(* IEC 61131-3 sources: JingjiangMoonbox/Application/Application/任务列表/Main_Task/IO配置表_1/KESAI1, 7 files *)

(* ---- KS_AbsEncModule_IODeal_KS1.st ---- *)
(*@CES
Name=KS_AbsEncModule_IODeal_KS1
Type=FunctionBlock
TypeGuid=6f9dac99-8de1-4efc-8465-68ac443b7d08
Guid=41d52946-2a11-4c79-a8c5-b68088c6a3a7
HasDeclaration=True
HasImplementation=False
*)
{DECLARATION}
FUNCTION_BLOCK KS_AbsEncModule_IODeal_KS1
VAR_INPUT
	i_xInputEn:BOOL;
	i_xOutPutEn:BOOL;
	(*这些值的处理未考虑双收双放*)
	i_pdwAbsEncSinglePos_Uw:POINTER TO DWORD;
	i_pwAbsEncMultiPos_Uw:POINTER TO WORD;
	(*收料*)
	i_pdwAbsEncSinglePos_Rw:POINTER TO DWORD;
	i_pwAbsEncMultiPos_Rw:POINTER TO WORD;
	//2025.08.20.152113+
	i_pstStAbsEncIOModule_Uw:POINTER TO StAbsEncIOModule;
	i_pstStAbsEncIOModule_Rw:POINTER TO StAbsEncIOModule;

END_VAR
VAR
	wIWTest:WORD;
	wQWTest: WORD;
	byAbsEncSts: BOOL;
END_VAR

{IMPLEMENTATION}

(* ---- KS_FB_IOMAP_AIAO_KS1.st ---- *)
(*@CES
Name=KS_FB_IOMAP_AIAO_KS1
Type=FunctionBlock
TypeGuid=6f9dac99-8de1-4efc-8465-68ac443b7d08
Guid=356f4cce-85a0-44c7-ab1e-a67fad378d86
HasDeclaration=True
HasImplementation=False
*)
{DECLARATION}
FUNCTION_BLOCK KS_FB_IOMAP_AIAO_KS1
VAR_INPUT
	i_xEn: BOOL;(*功能块使能|*)
	i_xRdInput: BOOL;(*读io输入|*)
	i_xWrOutput: BOOL;(*写io输出|*)
	i_pstStSysParam								: POINTER TO StSysParam;
	i_pastStProgMonitoring						: POINTER TO ARRAY [1..2] OF StProgMonitoring;
END_VAR
VAR_OUTPUT
	o_xEno: BOOL;(*indicated to i_xEn|*)
	o_iErNo: INT;(*0.no err\-1.bad parameter|*)
END_VAR
VAR
//	fb_KS_FB_SetAIType: KS_FB_SetAIType;
	fbKS_FB_Analog_IO_CTL: KS_FB_Analog_IO_CTL;

	byAiFilterTms_UwRw_I					:  BYTE:= 1;(*滤波次数*)
	byAiFilterTms_UwRw_II					:  BYTE:= 1;
	byAiFilterTms_IfOf_I					:  BYTE:= 1;
	byAiFilterTms_IfOf_II					:  BYTE:= 1;
	byAiFilterTms_DiaMeasure_I				:   BYTE:= 1;
	byAiFilterTms_DiaMeasure_II				:   BYTE:= 1;
END_VAR

{IMPLEMENTATION}

(* ---- KS_FB_IOMAP_Axis_KS1.st ---- *)
(*@CES
Name=KS_FB_IOMAP_Axis_KS1
Type=FunctionBlock
TypeGuid=6f9dac99-8de1-4efc-8465-68ac443b7d08
Guid=5e1ef807-2a8d-4def-8e48-4f55f608734d
HasDeclaration=True
HasImplementation=False
*)
{DECLARATION}
FUNCTION_BLOCK KS_FB_IOMAP_Axis_KS1
VAR_INPUT
	i_xEn: BOOL;(*功能块使能|*)
	i_xRdInput: BOOL;(*读io输入|*)
	i_xWrOutput: BOOL;(*写io输出|*)
	i_pastStIOMap_Axis_FE						: POINTER TO ARRAY [1..MAX_UNIT_NUM] OF StIOMap_Axis_FE;(*轴io数据区域|*)
END_VAR
VAR_OUTPUT
	o_xEno										: BOOL;(*indicated to i_xEn|*)
	o_iErNo										: INT;(*0.no err\-1.bad parameter|*)
END_VAR
VAR
	afbKS_FB_IOMap_Axis							: ARRAY [1..MAX_UNIT_NUM] OF KS_FB_MapAxisIOBasic;(*色组IO配置*)
END_VAR

{IMPLEMENTATION}

(* ---- KS_FB_IOMAP_AxisExtra_KS1.st ---- *)
(*@CES
Name=KS_FB_IOMAP_AxisExtra_KS1
Type=FunctionBlock
TypeGuid=6f9dac99-8de1-4efc-8465-68ac443b7d08
Guid=0dfac2a8-afaf-47de-8dd3-fd80962ebd90
HasDeclaration=True
HasImplementation=False
*)
{DECLARATION}
FUNCTION_BLOCK KS_FB_IOMAP_AxisExtra_KS1
VAR_INPUT
	i_xEn: BOOL;(*功能块使能|*)
	i_xRdInput: BOOL;(*读io输入|*)
	i_xWrOutput: BOOL;(*写io输出|*)
	i_pastStIOMap_Axis_Extra_FE						: POINTER TO ARRAY [1..MAX_UNIT_NUM] OF StIOMap_Axis_Extra_FE;(*轴io数据区域|*)
END_VAR
VAR_OUTPUT
	o_xEno										: BOOL;(*indicated to i_xEn|*)
	o_iErNo										: INT;(*0.no err\-1.bad parameter|*)
END_VAR
VAR
	afbKS_FB_IOMap_AxisExtra							: ARRAY [1..MAX_UNIT_NUM] OF KS_FB_MapAxisIOExtra;(*色组IO配置*)
END_VAR

{IMPLEMENTATION}

(* ---- KS_FB_IOMAP_Main_KS1.st ---- *)
(*@CES
Name=KS_FB_IOMAP_Main_KS1
Type=FunctionBlock
TypeGuid=6f9dac99-8de1-4efc-8465-68ac443b7d08
Guid=9ec1f607-9ce0-40a9-b7b7-7ca01d00a040
HasDeclaration=True
HasImplementation=False
*)
{DECLARATION}
FUNCTION_BLOCK KS_FB_IOMAP_Main_KS1
(*主面板IO配置分A/B系和放/收牵*)
(*正常单收单放选1和2*)
(*双收双放1和2是A系的放牵收牵，3和4是B系的放牵收牵*)
(*双收双放A放B收1和4*)
VAR_INPUT
	i_xEn: BOOL;(*功能块使能|*)
	i_xRdInput: BOOL;(*读io输入|*)
	i_xWrOutput: BOOL;(*写io输出|*)
	i_pastStIOMap_Main_FE						: POINTER TO ARRAY [1..4] OF StIOMap_Main_FE;(*轴io数据区域|*)
END_VAR
VAR_OUTPUT
	o_xEno										: BOOL;(*indicated to i_xEn|*)
	o_iErNo										: INT;(*0.no err\-1.bad parameter|*)
END_VAR
VAR
	afbKS_FB_MapIO_Main						: ARRAY [1..4] OF KS_FB_MapIO_Main;(*主面板IO配置*)
END_VAR

{IMPLEMENTATION}

(* ---- KS_FB_IOMAP_UwRw_KS1.st ---- *)
(*@CES
Name=KS_FB_IOMAP_UwRw_KS1
Type=FunctionBlock
TypeGuid=6f9dac99-8de1-4efc-8465-68ac443b7d08
Guid=3fdf527d-7ba2-4b44-94e3-31e35d6ee8ed
HasDeclaration=True
HasImplementation=False
*)
{DECLARATION}
 FUNCTION_BLOCK KS_FB_IOMAP_UwRw_KS1
VAR_INPUT
	i_xEn: BOOL;(*功能块使能|*)
	i_xRdInput: BOOL;(*读io输入|*)
	i_xWrOutput: BOOL;(*写io输出|*)
	i_pastStIOMap_UwRw_FE_Uw					: POINTER TO ARRAY [1..2] OF StIOMap_UwRw_FE;(*轴io数据区域|*)
	i_pastStIOMap_UwRw_FE_Rw					: POINTER TO ARRAY [1..2] OF StIOMap_UwRw_FE;(*轴io数据区域|*)
END_VAR
VAR_OUTPUT
	o_xEno										: BOOL;(*indicated to i_xEn|*)
	o_iErNo										: INT;(*0.no err\-1.bad parameter|*)
END_VAR
VAR
	afbKS_FB_MapIO_UwRw_Uw						: ARRAY [1..2] OF KS_FB_MapIO_UwRw;
	afbKS_FB_MapIO_UwRw_Rw						: ARRAY [1..2] OF KS_FB_MapIO_UwRw;
END_VAR

{IMPLEMENTATION}

(* ---- KS_FB_StepDriveIODeal_KS1.st ---- *)
(*@CES
Name=KS_FB_StepDriveIODeal_KS1
Type=FunctionBlock
TypeGuid=6f9dac99-8de1-4efc-8465-68ac443b7d08
Guid=61a728a1-12ea-4f97-af25-7b7b77ea73c8
HasDeclaration=True
HasImplementation=False
*)
{DECLARATION}
FUNCTION_BLOCK KS_FB_StepDriveIODeal_KS1
VAR_INPUT
	i_xInputEn:BOOL;
	i_xOutPutEn:BOOL;
	i_pastStDigitalMicroStepDrive :POINTER TO  ARRAY [1..MAX_UNIT_NUM] OF StDigitalMicroStepDrive;
	i_pastStStepDriveIOModule:POINTER TO ARRAY [1..MAX_UNIT_NUM] OF StStepDriveIOModule;
	i_pastStEnc0410R:POINTER TO ARRAY [1..MAX_UNIT_NUM] OF StEnc0410R;
END_VAR
VAR_OUTPUT
END_VAR
VAR
	wTest: WORD;
	afbKS_FB_StepDriveIOModule: ARRAY [1..MAX_UNIT_NUM] OF KS_FB_StepDriveIOModule;
END_VAR

{IMPLEMENTATION}
